Fanuc KAREL source: kc00019.KL

-- PROVISIONAL review KL for V1013-1; original PC SHA256 5b20b916a1245567c6a3e519b3262274136493a0835c8b46e4362909c291e6d1
-- Incomplete behavior may be omitted. Consult companion uncertainty JSON. Do not deploy.
PROGRAM KC00019
%NOLOCKGROUP
BEGIN
  -- UNRESOLVED_PC offsets 5-53; opcodes 27,22,22,22,22,22,2A,22,22,31
  -- UNRESOLVED_PC offsets 58-62; opcodes 7F
END KC00019
